(* IEC 61131-3 sources: Elmo_Master/Lasal_PRG/Elmo_EtherCAT_Test_4Axis/Class/SafetyManager (part 6) *)

      UdpReceiveData.SectionStop();
    else
      //sequence counter is not the same
      sUdpVars.WrongSequenceInResponseCnt += 1;

      //check the sequence difference, it could be a retry from other side which contains sdo data
      SequenceDifference := pConnection^.ActReceiveData.udSequenceNumber$DINT - pConnection^.ActSendData.udSequenceNumber$DINT;

      UdpReceiveData.SectionStart();
      //if Sequence difference is -1 it could be a response retry with sdo data
      if (pPacket^.Header.SdoDataLength) & (pConnection^.ActReceiveData.SdoLength = 0)
      & (pPacket^.Header.SdoDataLength <= UDP_MAX_SDO_SIZE) & (SequenceDifference = -1) then
        pConnection^.ActReceiveData.SdoLength := pPacket^.Header.SdoDataLength;
        _memcpy(ptr1:=#pConnection^.ActReceiveData.SdoData, ptr2:=#pPacket^.Data + pConnection^.ActReceiveData.PdoLength, cntr:=pConnection^.ActReceiveData.SdoLength);
      end_if;
      UdpReceiveData.SectionStop();
    end_if;

    // save safety number of other side
    pConnection^.SafetyNbrOtherSide       := pPacket^.Header.SafetyNbr;
  else
    sUdpVars.WrongReceiveUDPLength += 1;
  end_if;

END_FUNCTION

FUNCTION SafetyManager::ForwardReceivedUdpSDOs
  VAR_INPUT
    paConnections 	: ^t_aUdpConnections;
    ConnectionNo 	: UDINT;
  END_VAR
  VAR
    i               : UDINT;
    pActConnection  : ^t_UdpConnection;
    pHelpCfg        : ^t_CfgListElem;
    pHelpModule     : ^t_ModuleListElem;
    InterfaceCRC    : HDINT;
    SafetyNumber    : HDINT;
    MyPara          : CmdStruct;
    MyResult        : results;
    pDO 	          : ^SafetyCDIAS_Base::SDOHeader;
    pCompDestPath   : ^USINT;
    pHelpSafety     : ^t_SafetyComponent;
    ResponseValue   : BOOL;
    FoundTarget     : BOOL;
  END_VAR

  ResponseValue := paConnections = sUdpVars.paConnectionsToProducers;

  pActConnection := #paConnections^[0];
  for i := 0 to (ConnectionNo-1) do

    // check if there is a SDO to forward
    if pActConnection^.ActReceiveData.SdoLength then

      FoundTarget := FALSE;

      UdpReceiveData.SectionStart();

      // get a pointer to the compressed destination path
      pDO := (#pActConnection^.ActReceiveData.SdoData)$^SafetyCDIAS_Base::SDOHeader;
      if (pDO^.StdHeader.Typ.Response = ResponseValue) then
        pCompDestPath := (#pDO^.DstAdr)$^USINT;

        // check if it's addressed by topology path and it's an IP
        if ((pDO^.StdHeader.Typ AND SSDO_MASK_TYPE) = FRM_TYPECODE_SSDO_MOD_TP) & (pCompDestPath^ = INTERFACE_IP_MODE) then
          // after the mode byte we find the interface CRC
          InterfaceCRC := ((pCompDestPath + 1)$^HDINT)^;

          // search all configs, all moduleconfigs

          pHelpCfg := pConfigs;
          while pHelpCfg & pActConnection^.ActReceiveData.SdoLength do
            pHelpModule := pHelpCfg^.pFirstModuleCfg;
            while pHelpModule & pActConnection^.ActReceiveData.SdoLength do
              if pHelpModule^.ModuleInfo.InterfaceCRC = InterfaceCRC then
                // we found the interface CRC, now we have to make a connection via the SafetyNumber between the actual module config and the module handles
                pHelpSafety := pFirstSafetyComponent;
                while pHelpSafety & pActConnection^.ActReceiveData.SdoLength do
                  // we compare the safety number
                  if pHelpSafety^.SafetyNbr = pHelpModule^.ModuleInfo.SafetyNbr then

                    MyPara.uiCmd := CMD_SM_SDO_TO_MODULE;
                    MyPara.aPara[0] := pActConnection^.ActReceiveData.SdoLength;
                    MyPara.aPara[1] := (#pActConnection^.ActReceiveData.SdoData)$DINT;
                    MyPara.aPara[2] := this$DINT;

                    pHelpSafety^.pThis^.NewInst(#MyPara, #MyResult);

                    FoundTarget := TRUE;
                  end_if;

                  pHelpSafety := pHelpSafety^.pNext;
                end_while;
              end_if;

              pHelpModule := pHelpModule^.pNext;
            end_while;

            pHelpCfg := pHelpCfg^.pNext;
          end_while;
        else
          SafetyNumber := pDO^.DstAdr;

          // search by safety number and forward to internal module
          pHelpSafety := pFirstSafetyComponent;
          while pHelpSafety & pActConnection^.ActReceiveData.SdoLength do
            // we compare the safety number
            if pHelpSafety^.SafetyNbr = SafetyNumber then
              MyPara.uiCmd := CMD_SM_SDO_TO_MODULE;
              MyPara.aPara[0] := pActConnection^.ActReceiveData.SdoLength;
              MyPara.aPara[1] := (#pActConnection^.ActReceiveData.SdoData)$DINT;
              MyPara.aPara[2] := this$DINT;

              pHelpSafety^.pThis^.NewInst(#MyPara, #MyResult);

              FoundTarget := TRUE;
            end_if;

            pHelpSafety := pHelpSafety^.pNext;
          end_while;
        end_if;

        // reset length if the response bit matches (if we found it, we already forwarded it. if not, we're not going to find it next time)
        pActConnection^.ActReceiveData.SdoLength := 0;
      else
        // check which list it is
        if ResponseValue then
          sUdpVars.InvalidResponseSettingAtFowardingProducerList += 1;
        else
          sUdpVars.InvalidResponseSettingAtFowardingConsumerList += 1;
        end_if;
      end_if;

      UdpReceiveData.SectionStop();

    end_if;

    pActConnection += sizeof(t_UdpConnection);
  end_for;

END_FUNCTION

FUNCTION SafetyManager::ForwardSDO2UdpBySafetyNbr
  VAR_INPUT
    SDOLength 	: UINT;
    pSDO 	: ^USINT;
  END_VAR
  VAR_OUTPUT
    FoundTarged 	: BOOL;
  END_VAR
  VAR
    i               : UDINT;
    pActConnection  : ^t_UdpConnection;
    TargetSafetyNbr : HDINT;
    pDO 	          : ^SafetyCDIAS_Base::SDOHeader;
  END_VAR

  FoundTarged := FALSE;

  // get a pointer to the compressed destination path
  pDO := pSDO$^SafetyCDIAS_Base::SDOHeader;
  TargetSafetyNbr := pDO^.DstAdr;

  if sUdpVars.ConsumerConnectionNo then
    pActConnection := #sUdpVars.paConnectionsToConsumers^[0];
    for i := 0 to (sUdpVars.ConsumerConnectionNo-1) do
      // the safety number has to match and since it's a message to a consumer it has to be a response
      if (pActConnection^.SafetyNbrOtherSide = TargetSafetyNbr) & (pDO^.StdHeader.Typ.Response = TRUE) then
        // got it => forward the SDO
        if SDOLength <= UDP_MAX_SDO_SIZE then
          // check for unsent SDO first
          if pActConnection^.ActSendData.SdoLength = 0 then
            UdpSendData.SectionStart();

            _memcpy(ptr1:=#pActConnection^.ActSendData.SdoData, ptr2:=pSDO, cntr:=SDOLength);
            pActConnection^.ActSendData.SdoLength     := SDOLength$USINT;

            UdpSendData.SectionStop();
          else
            sUdpVars.SdoAlreadyUsedCnt += 1;
          end_if;
        else
          LogError("@046E (SafetyManager::ForwardSDO2UdpBySafetyNbr) SDO size exceeds the allowed size (Compressed Topology Path: UDP)");
        end_if;

        FoundTarged := TRUE;
        return;
      end_if;

      pActConnection += sizeof(t_UdpConnection);
    end_for;
  end_if;

  if sUdpVars.ProducerConnectionNo then
    pActConnection := #sUdpVars.paConnectionsToProducers^[0];
    for i := 0 to (sUdpVars.ProducerConnectionNo-1) do
      // the safety number has to match and since it's a message to a producer it has to be a request
      if (pActConnection^.SafetyNbrOtherSide = TargetSafetyNbr) & (pDO^.StdHeader.Typ.Response = FALSE) then
        // got it => forward the SDO
        if SDOLength <= UDP_MAX_SDO_SIZE then
          // check for unsent SDO first
          if pActConnection^.ActSendData.SdoLength = 0 then
            UdpSendData.SectionStart();

            _memcpy(ptr1:=#pActConnection^.ActSendData.SdoData, ptr2:=pSDO, cntr:=SDOLength);
            pActConnection^.ActSendData.SdoLength     := SDOLength$USINT;

            UdpSendData.SectionStop();
          else
            sUdpVars.SdoAlreadyUsedCnt += 1;
          end_if;
        else
          LogError("@046E (SafetyManager::ForwardSDO2Udp) SDO size exceeds the allowed size (Compressed Topology Path: UDP)");
        end_if;

        FoundTarged := TRUE;
        return;
      end_if;

      pActConnection += sizeof(t_UdpConnection);
    end_for;
  end_if;

END_FUNCTION

FUNCTION SafetyManager::ShareUdpConnectionInfos
  VAR
    i                 : UDINT;
    pUdpConnection    : ^t_UdpConnection;
    AnythingMissing   : BOOL;
    ActInitialized    : BOOL;
    FoundConnection   : BOOL;
    pHelpSafety       : ^t_SafetyComponent;
    pHelpCfg          : ^t_CfgListElem;
    pFSoEConnection   : ^t_FSoEConnectionDetails;
    MyPara            : CmdStruct;
    MyResult          : results;
    retcode           : iprStates;

    ModuleReadOffset  : UINT;
    ModuleReadSize    : UINT;
    ModuleWriteOffset : UINT;
    ModuleWriteSize   : UINT;
    MngReadOffset     : UINT;
    MngReadSize       : UINT;
    MngWriteOffset    : UINT;
    MngWriteSize      : UINT;
  END_VAR

  AnythingMissing := FALSE;

  if sUdpVars.ConsumerConnectionNo then
    pUdpConnection := #sUdpVars.paConnectionsToConsumers^[0];
    for i := 0 to (sUdpVars.ConsumerConnectionNo-1) do
      // check if we received something so far at this connection
      if (pUdpConnection^.ReceivedPackages & (pUdpConnection^.InfoBits.PdosInitialized = FALSE)) then
        FoundConnection := ActInitialized := FALSE;

        // check FSoE Connections in the available configs if there is a match at the interface CRC
        pHelpCfg := pConfigs;
        while pHelpCfg & (FoundConnection = FALSE) do
          pFSoEConnection := pHelpCfg^.pFirstFSoEConnection;
          while pFSoEConnection & (FoundConnection = FALSE) do
            // only interface slave connections which are not used yet are relevant
            if pFSoEConnection^.Flags.IsInterfaceConnection & (pFSoEConnection^.Flags.IsMaster = FALSE) & (pFSoEConnection^.InternalConnectionState = FCS_RESET) &
               pFSoEConnection^.pSlavePathComp & ((pFSoEConnection^.pSlavePathComp$^HDINT + 1)^ = pUdpConnection^.IFCRC) then

              // found the connection
              FoundConnection := TRUE;

              // now try to initialize it

              pHelpSafety := pFirstSafetyComponent;
              while pHelpSafety do
                if pHelpSafety^.SafetyNbr = pFSoEConnection^.OwnerSafetyNbr then
                  exit;
                end_if;

                pHelpSafety := pHelpSafety^.pNext;
              end_while;

              if pHelpSafety then
#ifdef SAFETY_DEBUG_LOGGING_ACTIVATED
#pragma message("RamAnd 20.11.2014 16:41 \ testweise mapping loggen")
                LogValue("@DBG (SafetyManager::ShareUdpConnectionInfos) <This side is Slave> ConnectionID: 0x{0}, SlaveAddress: 0x{1}, IFCRC: 0x{2}", Value:=pFSoEConnection^.ConnectionID, Value2:=pFSoEConnection^.SlaveAddress, Value3 := (pFSoEConnection^.pSlavePathComp$^HDINT + 1)^);
                LogValue("@DBG (SafetyManager::ShareUdpConnectionInfos) <This side is Slave> UdpInfo: SNr: 0x{0}, SNrOtherSide: 0x{1}, IFCRC: 0x{2}", Value:=pUdpConnection^.SafetyNbr, Value2:=pUdpConnection^.SafetyNbrOtherSide, Value3 := pUdpConnection^.IFCRC);
#endif

                // the module is slave and the managing module master
                ModuleReadOffset  := pFSoEConnection^.SlaveReadOffset;
                ModuleReadSize    := pFSoEConnection^.MasterWriteSize;
                ModuleWriteOffset := pFSoEConnection^.SlaveWriteOffset;
                ModuleWriteSize   := pFSoEConnection^.MasterReadSize;
                MngReadOffset     := 0; // offsets in managing modules are always dynamic
                MngReadSize       := pFSoEConnection^.MasterReadSize;
                MngWriteOffset    := 0; // offsets in managing modules are always dynamic
                MngWriteSize      := pFSoEConnection^.MasterWriteSize;

#ifdef SAFETY_DEBUG_LOGGING_ACTIVATED
#pragma message("RamAnd 20.11.2014 16:41 \ testweise mapping loggen")
                LogValue("@DBG (SafetyManager::ShareUdpConnectionInfos) Modul => Udp: Rd Offset Modul: 0x{0}, IP: 0x{1}, Größe: 0x{2}", Value:=ModuleReadOffset, Value2:=pUdpConnection^.IP, Value3:=ModuleReadSize);
#endif

                MyPara.uiCmd    := CMD_SM_ADD_INPUT_PDO;
                MyPara.aPara[0] := (#pUdpConnection^.ThreadSafePdoReceiveBuffer)$DINT;
                MyPara.aPara[1] := 0;
                MyPara.aPara[2] := pUdpConnection^.SafetyNbrOtherSide$DINT;
                MyPara.aPara[3] := ModuleWriteSize;
                MyPara.aPara[4] := 0;
                MyPara.aPara[5] := 0;
                MyPara.aPara[6] := 0;
                MyPara.aPara[7] := ModuleWriteOffset;
                MyPara.aPara[8] := SM_IF_VALIDITY_MARK$DINT;
                MyPara.aPara[9] := TRUE;

                retcode := pHelpSafety^.pThis^.NewInst(#MyPara, #MyResult);

                if retcode = ERROR then
                  LogError("@0848 (SafetyManager::ShareUdpConnectionInfos) Failed to add input PDO for a connection to a Consumer");

                  // mark the connection to not try again later
                  pFSoEConnection^.InternalConnectionState := FCS_NOT_INITIALIZED;

                  return;
                elsif retcode = BUSY then
                  // try again later (skip further initialisation steps)
                  return;
                end_if;

                if FSoEInputPDONo < MAX_FSOE_CONNECTIONS then
                  aFSoEInputPDOs[FSoEInputPDONo].pSafety    := pHelpSafety;
                  aFSoEInputPDOs[FSoEInputPDONo].pMem       := MyPara.aPara[0];
                  FSoEInputPDONo                            += 1;

                  pUdpConnection^.ActReceiveData.PdoLength  := ModuleWriteSize;
                else
                  LogValue("@0490 (SafetyManager::ShareUdpConnectionInfos) Maximum limit of allowed FSoE input Frames exceeded (0x{0})", Value:=MAX_FSOE_CONNECTIONS);
                  exit;
                end_if;

                if sUdpVars.ReceiveCopyCmdNo < MAX_UDP_IF_ALLOWED then
                  sUdpVars.aReceiveCopyCmds[sUdpVars.ReceiveCopyCmdNo].pSource      := (#pUdpConnection^.ActReceiveData.PdoData)$^USINT;
                  sUdpVars.aReceiveCopyCmds[sUdpVars.ReceiveCopyCmdNo].pDest        := MyPara.aPara[0]$^USINT;
                  sUdpVars.aReceiveCopyCmds[sUdpVars.ReceiveCopyCmdNo].Size         := ModuleWriteSize;
                  sUdpVars.ReceiveCopyCmdNo                                            += 1;
                else
                  LogValue("@049F (SafetyManager::ShareUdpConnectionInfos) Maximum limit of allowed UDP receive copy commands exceeded (0x{0})", Value:=MAX_UDP_IF_ALLOWED);
                  exit;
                end_if;

                MyPara.uiCmd    := CMD_SM_ADD_OUTPUT_PDO;
                MyPara.aPara[0] := 1;  // mark as interface frame PDO
                pHelpSafety^.pThis^.NewInst(#MyPara, #MyResult);

//                  pPDOElement^.SourceInfo.pPDOMem       := MyResult.aData[0]$^USINT;
//                  pPDOElement^.SourceInfo.pPDOMemDPRAM  := MyResult.aData[4]$^USINT;
//                  pPDOElement^.SourceInfo.HandlePDODPRAM:= MyResult.aData[8]$UDINT;   // Needed for Payload Support
//                  pPDOElement^.SourceInfo.OffsetPDODPRAM:= MyResult.aData[12]$UDINT;  // Needed for Payload Support

                if sUdpVars.SendCopyCmdNo < MAX_UDP_IF_ALLOWED then
                  sUdpVars.aSendCopyCmds[sUdpVars.SendCopyCmdNo].pSource      := MyResult.aData[0]$^USINT + ModuleReadOffset;
                  sUdpVars.aSendCopyCmds[sUdpVars.SendCopyCmdNo].pDest        := #pUdpConnection^.ActSendData.PdoData;
                  sUdpVars.aSendCopyCmds[sUdpVars.SendCopyCmdNo].Size         := ModuleReadSize;
                  sUdpVars.SendCopyCmdNo                                         += 1;

                  pUdpConnection^.ActSendData.PdoLength           := ModuleReadSize;
                else
                  LogValue("@049E (SafetyManager::ShareUdpConnectionInfos) Maximum limit of allowed UDP send copy commands exceeded (0x{0})", Value:=MAX_UDP_IF_ALLOWED);
                  exit;
                end_if;

#ifdef SAFETY_DEBUG_LOGGING_ACTIVATED
#pragma message("RamAnd 20.11.2014 16:41 \ testweise mapping loggen")
                LogValue("@DBG (SafetyManager::ShareUdpConnectionInfos) Udp => Modul: Wr Offset Modul: 0x{0}, IP: 0x{1}, Größe: 0x{2}", Value:=ModuleWriteOffset, Value2:=pUdpConnection^.IP, Value3:=ModuleWriteSize);
#endif

                // mark the FSoE connection as established
                pFSoEConnection^.InternalConnectionState  := FCS_CONNECTION;

                // mark the udp connection as established
                pUdpConnection^.InfoBits.PdosInitialized  := TRUE;

                // connection initialized
                ActInitialized                            := TRUE;

                // check if we have all slave addresses now
                CheckLocalSlaveAddresses();
              else
                LogValue("@495 (SafetyManager::ShareUdpConnectionInfos) Could not find safety module with safety number 0x{0} for FSoE interface connection", Value:=pFSoEConnection^.OwnerSafetyNbr);
              end_if;
            end_if;

            pFSoEConnection := pFSoEConnection^.pNext;
          end_while;

          if pHelpCfg then
            pHelpCfg := pHelpCfg^.pNext;
          end_if;
        end_while;

        if ActInitialized = FALSE then
          AnythingMissing := TRUE;
        end_if;
      elsif (pUdpConnection^.ReceivedPackages = 0) then
        AnythingMissing := TRUE;
      end_if;

      pUdpConnection += sizeof(t_UdpConnection);
    end_for;
  end_if;

  if sUdpVars.ProducerConnectionNo then
    pUdpConnection := #sUdpVars.paConnectionsToProducers^[0];
    for i := 0 to (sUdpVars.ProducerConnectionNo-1) do
      // check if we received something so far at this connection
      if (pUdpConnection^.ReceivedPackages & (pUdpConnection^.InfoBits.PdosInitialized = FALSE)) then
        FoundConnection := ActInitialized := FALSE;

        // check FSoE Connections in the available configs if there is a match at the interface CRC
        pHelpCfg := pConfigs;
        while pHelpCfg & (FoundConnection = FALSE) do
          pFSoEConnection := pHelpCfg^.pFirstFSoEConnection;
          while pFSoEConnection & (FoundConnection = FALSE) do
            // only interface master connections which are not used are relevant
            if pFSoEConnection^.Flags.IsInterfaceConnection & pFSoEConnection^.Flags.IsMaster & (pFSoEConnection^.InternalConnectionState = FCS_RESET) then
              // check if it's our connection
              if ( pFSoEConnection^.pSlavePathComp) &
                 ( pFSoEConnection^.pSlavePathComp^             = INTERFACE_IP_MODE) &
                 ((pFSoEConnection^.pSlavePathComp$^HDINT + 1)^ = pUdpConnection^.IFCRC) &
                 ((pFSoEConnection^.pSlavePathComp$^HDINT + 5)^ = pUdpConnection^.IP) then

                // found the connection
                FoundConnection := TRUE;

                // now try to initialize it

                pHelpSafety := pFirstSafetyComponent;
                while pHelpSafety do
                  if pHelpSafety^.SafetyNbr = pFSoEConnection^.OwnerSafetyNbr then
                    exit;
                  end_if;

                  pHelpSafety := pHelpSafety^.pNext;
                end_while;

                if pHelpSafety then
  #ifdef SAFETY_DEBUG_LOGGING_ACTIVATED
  #pragma message("RamAnd 20.11.2014 16:41 \ testweise mapping loggen")
                  LogValue("@DBG (SafetyManager::ShareUdpConnectionInfos) <This side is Master> ConnectionID: 0x{0}, SlaveAddress: 0x{1}, InterfaceCRC: 0x{2}", Value:=pFSoEConnection^.ConnectionID, Value2:=pFSoEConnection^.SlaveAddress, Value3 := pUdpConnection^.IFCRC);
#endif

                  // the module is master and the managing module slave
                  ModuleReadOffset  := pFSoEConnection^.MasterReadOffset;
                  ModuleReadSize    := pFSoEConnection^.MasterReadSize;
                  ModuleWriteOffset := pFSoEConnection^.MasterWriteOffset;
                  ModuleWriteSize   := pFSoEConnection^.MasterWriteSize;
                  MngReadOffset     := 0; // offsets in managing modules are always dynamic
                  MngReadSize       := pFSoEConnection^.MasterWriteSize;
                  MngWriteOffset    := 0; // offsets in managing modules are always dynamic
                  MngWriteSize      := pFSoEConnection^.MasterReadSize;

  #ifdef SAFETY_DEBUG_LOGGING_ACTIVATED
  #pragma message("RamAnd 20.11.2014 16:41 \ testweise mapping loggen")
                  LogValue("@DBG (SafetyManager::ShareUdpConnectionInfos) Modul => Udp: Rd Offset Modul: 0x{0}, IP: 0x{1}, Größe: 0x{2}", Value:=ModuleReadOffset, Value2:=pUdpConnection^.IP, Value3:=ModuleReadSize);
  #endif

                  MyPara.uiCmd    := CMD_SM_ADD_INPUT_PDO;
                  MyPara.aPara[0] := (#pUdpConnection^.ThreadSafePdoReceiveBuffer)$DINT;
                  MyPara.aPara[1] := 0;
                  MyPara.aPara[2] := pUdpConnection^.SafetyNbrOtherSide$DINT;
                  MyPara.aPara[3] := ModuleWriteSize;
                  MyPara.aPara[4] := 0;
                  MyPara.aPara[5] := 0;
                  MyPara.aPara[6] := 0;
                  MyPara.aPara[7] := ModuleWriteOffset;
                  MyPara.aPara[8] := SM_IF_VALIDITY_MARK$DINT;
                  MyPara.aPara[9] := TRUE;

                  retcode := pHelpSafety^.pThis^.NewInst(#MyPara, #MyResult);

                  if retcode = ERROR then
                    LogError("@0849 (SafetyManager::ShareUdpConnectionInfos) Failed to add input PDO for a connection to a Producer");

                    // mark the connection to not try again later
                    pFSoEConnection^.InternalConnectionState := FCS_NOT_INITIALIZED;

                    return;
                  elsif retcode = BUSY then
                    // try again later (skip further initialisation steps)
                    return;
                  end_if;

                  if FSoEInputPDONo < MAX_FSOE_CONNECTIONS then
                    aFSoEInputPDOs[FSoEInputPDONo].pSafety    := pHelpSafety;
                    aFSoEInputPDOs[FSoEInputPDONo].pMem       := MyPara.aPara[0];
                    FSoEInputPDONo += 1;

                    pUdpConnection^.ActReceiveData.PdoLength  := ModuleWriteSize;
                  else
                    LogValue("@0490 (SafetyManager::ShareUdpConnectionInfos) Maximum limit of allowed FSoE input Frames exceeded (0x{0})", Value:=MAX_FSOE_CONNECTIONS);
                    exit;
                  end_if;

                  if sUdpVars.ReceiveCopyCmdNo < MAX_UDP_IF_ALLOWED then
                    sUdpVars.aReceiveCopyCmds[sUdpVars.ReceiveCopyCmdNo].pSource  := (#pUdpConnection^.ActReceiveData.PdoData)$^USINT;
                    sUdpVars.aReceiveCopyCmds[sUdpVars.ReceiveCopyCmdNo].pDest    := MyPara.aPara[0]$^USINT;
                    sUdpVars.aReceiveCopyCmds[sUdpVars.ReceiveCopyCmdNo].Size     := ModuleWriteSize;
                    sUdpVars.ReceiveCopyCmdNo                                        += 1;
                  else
                    LogValue("@049F (SafetyManager::ShareUdpConnectionInfos) Maximum limit of allowed UDP receive copy commands exceeded (0x{0})", Value:=MAX_UDP_IF_ALLOWED);
                    exit;
                  end_if;

                  MyPara.uiCmd      := CMD_SM_ADD_OUTPUT_PDO;
                  MyPara.aPara[0]   := 1;  // mark as interface frame PDO
                  pHelpSafety^.pThis^.NewInst(#MyPara, #MyResult);

  //                  pPDOElement^.SourceInfo.pPDOMem       := MyResult.aData[0]$^USINT;
  //                  pPDOElement^.SourceInfo.pPDOMemDPRAM  := MyResult.aData[4]$^USINT;
  //                  pPDOElement^.SourceInfo.HandlePDODPRAM:= MyResult.aData[8]$UDINT;   // Needed for Payload Support
  //                  pPDOElement^.SourceInfo.OffsetPDODPRAM:= MyResult.aData[12]$UDINT;  // Needed for Payload Support

                  if sUdpVars.SendCopyCmdNo < MAX_UDP_IF_ALLOWED then
                    sUdpVars.aSendCopyCmds[sUdpVars.SendCopyCmdNo].pSource      := MyResult.aData[0]$^USINT + ModuleReadOffset;
                    sUdpVars.aSendCopyCmds[sUdpVars.SendCopyCmdNo].pDest        := #pUdpConnection^.ActSendData.PdoData;
                    sUdpVars.aSendCopyCmds[sUdpVars.SendCopyCmdNo].Size         := ModuleReadSize;
                    sUdpVars.SendCopyCmdNo                                         += 1;

                    pUdpConnection^.ActSendData.PdoLength                             := ModuleReadSize;
                  else
                    LogValue("@049E (SafetyManager::ShareUdpConnectionInfos) Maximum limit of allowed UDP send copy commands exceeded (0x{0})", Value:=MAX_UDP_IF_ALLOWED);
                    exit;
                  end_if;

  #ifdef SAFETY_DEBUG_LOGGING_ACTIVATED
  #pragma message("RamAnd 20.11.2014 16:41 \ testweise mapping loggen")
                  LogValue("@DBG (SafetyManager::ShareUdpConnectionInfos) Udp => Modul: Wr Offset Modul: 0x{0}, IP: 0x{1}, Größe: 0x{2}", Value:=ModuleWriteOffset, Value2:=pUdpConnection^.IP, Value3:=ModuleWriteSize);
  #endif

                  // mark the FSoE connection as established
                  pFSoEConnection^.InternalConnectionState  := FCS_CONNECTION;

                  // mark the udp connection as established
                  pUdpConnection^.InfoBits.PdosInitialized  := TRUE;

                  // connection initialized
                  ActInitialized                            := TRUE;

                  // check if we have all slave addresses now
                  CheckLocalSlaveAddresses();
                else
                  LogValue("@0495 (SafetyManager::ShareUdpConnectionInfos) Could not find safety module with safety number 0x{0} for FSoE interface connection", Value:=pFSoEConnection^.OwnerSafetyNbr);
                end_if;

              end_if;

            end_if;

            pFSoEConnection := pFSoEConnection^.pNext;
          end_while;

          pHelpCfg := pHelpCfg^.pNext;
       end_while;

        if ActInitialized = FALSE then
          AnythingMissing := TRUE;
        end_if;
      elsif (pUdpConnection^.ReceivedPackages = 0) then
        AnythingMissing := TRUE;
      end_if;

      pUdpConnection += sizeof(t_UdpConnection);
    end_for;
  end_if;

  // if all available udp connections are initialized => set the marker for not coming here any more
  if AnythingMissing = FALSE then
    sUdpVars.ConnectionsInitialized := TRUE;

    // update scheduler grid
    SetUdpSchedulerGrid();
  end_if;

END_FUNCTION

FUNCTION SafetyManager::SetUdpSchedulerGrid
  VAR
    Temp            : UDINT;
    bGetRequestTimeout : BOOL;
  END_VAR

  bGetRequestTimeout := FALSE;

  // we can only calculate if there are producer connections => otherwise the scheduler is not active
  if sUdpVars.ProducerConnectionNo then

    // the timeout is calculated so we could fit 4 timed out transmissions into the watchdog time (watchdog = 2*transmission time)
    Temp := sUdpVars.LowestTransmissionTime_ms * 2 / 4;

    // if the result is smaller than the minimum timeout => set it to the minimum
    if Temp < UDP_MIN_REQUEST_TIMEOUT then
      Temp := UDP_MIN_REQUEST_TIMEOUT;
    end_if;

    sUdpVars.CalculatedRequestTimeout := Temp;
    bGetRequestTimeout := TRUE;
  else
    // activate the default settings (min settings)
    sUdpVars.CalculatedRequestTimeout := UDP_MIN_REQUEST_TIMEOUT;
  end_if;

  // use default value for request time
  sUdpVars.CalculatedRequestTime    := UDP_MIN_REQUEST_TIME;

  //check for advanced request time from user
  if sUdpVars.udAdvancedRequestCycle >= UDP_MIN_REQUEST_TIME
  & sUdpVars.udAdvancedRequestCycle <= (sUdpVars.CalculatedRequestTimeout/2)  then
    sUdpVars.CalculatedRequestTime := sUdpVars.udAdvancedRequestCycle;
  else
    //only log error if we got calculated request timeout and value is not zero
    if bGetRequestTimeout = TRUE & sUdpVars.udAdvancedResponseTimeout <> 0 & bd_SingleLog.SetUdpRequestCycleFailed = FALSE then
      LogValue("@04D6 (SafetyManager::SetUdpSchedulerGrid) [SL] The value of 0x{0} for the UDP Request Cycle is not valid! The maximum value is 0x{1}", Value:=sUdpVars.udAdvancedRequestCycle, (sUdpVars.CalculatedRequestTimeout/2));
      bd_SingleLog.SetUdpRequestCycleFailed := TRUE;
    end_if;
  end_if;

  // always use the min settings for the responses
  sUdpVars.CalculatedResponseTime    := UDP_MIN_RESPONSE_TIME;
  sUdpVars.CalculatedResponseTimeout := UDP_MIN_RESPONSE_TIMEOUT;

  //check for advanced response timeout from user
  if sUdpVars.udAdvancedResponseTimeout >= UDP_MIN_RESPONSE_TIMEOUT then
    sUdpVars.CalculatedResponseTimeout := sUdpVars.udAdvancedResponseTimeout;
  else
    // only log error if value is not zero
    if sUdpVars.udAdvancedResponseTimeout <> 0 & bd_SingleLog.SetUdpResponseTimeoutFailed = FALSE then
      LogValue("@04D7 (SafetyManager::SetUdpSchedulerGrid) [SL] The value of 0x{0} for the UDP Response Timeout is not valid! The minimum value is 0x{1}", Value:=sUdpVars.udAdvancedResponseTimeout, UDP_MIN_RESPONSE_TIMEOUT);
      bd_SingleLog.SetUdpResponseTimeoutFailed := TRUE;
    end_if;
  end_if;

  // if the override values are set => activate them here to override all other settings
  if sUdpVars.udOverrideCycleTime then
    // set the scheduler grid for requests and resonses according to the override value
    sUdpVars.CalculatedRequestTime  := sUdpVars.udOverrideCycleTime;
    sUdpVars.CalculatedResponseTime := sUdpVars.udOverrideCycleTime;
  end_if;

  if sUdpVars.udOverrideTimeout then
    // set the timeout value for requests and resonses according to the override value
    sUdpVars.CalculatedRequestTimeout  := sUdpVars.udOverrideTimeout;
    sUdpVars.CalculatedResponseTimeout := sUdpVars.udOverrideTimeout;
  end_if;

END_FUNCTION

FUNCTION SafetyManager::UdpResponseScheduler
  VAR
    pActResponseEntry : ^t_UdpConnection;
    pActRetryEntry    : ^t_UdpConnection;
    tmpretcode        : DINT;
    i                 : UDINT;
  END_VAR

  //point to actual request-entry
  pActResponseEntry := #sUdpVars.paConnectionsToConsumers^[sUdpVars.ResponseScheduler.ActRequestedIndex];

  //send a request every TRequestTime x Cycnt Cycle
  if ((sUdpVars.ResponseScheduler.CyCnt MOD sUdpVars.CalculatedResponseTime) = 0) then

    // search through the list if something has to be sent (check also for changes in the data)
    for i := 0 to sUdpVars.ConsumerConnectionNo-1 do

      //only send a request if not waiting for a response and the IP is valid (on cleaning out the connections some may be set to 0)
      if (pActResponseEntry^.WaitForResponse = FALSE) & (pActResponseEntry^.IP <> 0) & (pActResponseEntry^.SendResponse = TRUE) then

        //send request to mover of actual entry
        tmpretcode := SendUdpResponse(pActResponseEntry);
        if tmpretcode >= 0 then

          //if sending was successful we are waiting for a response
          pActResponseEntry^.WaitForResponse := TRUE;
          pActResponseEntry^.SendResponse    := FALSE;
          pActResponseEntry^.TLastRequest      := ops.tAbsolute;
          pActResponseEntry^.RequestRetries    := 0;

        else
          //unable to send request
          if bd_SingleLog.SendUdpRspFailed = FALSE then
            bd_SingleLog.SendUdpRspFailed := TRUE;
            LogError("@04A0 (SafetyManager::UdpResponseScheduler) [SL] Failed to send udp response");
          end_if;
        end_if;

      end_if;

      //increase actual index
      if sUdpVars.ResponseScheduler.ActRequestedIndex < (sUdpVars.ConsumerConnectionNo-1) then
        sUdpVars.ResponseScheduler.ActRequestedIndex += 1;
      else
        //when reaching last entry -> reset index
        sUdpVars.ResponseScheduler.ActRequestedIndex := 0;
      end_if;

      pActResponseEntry := #sUdpVars.paConnectionsToConsumers^[sUdpVars.ResponseScheduler.ActRequestedIndex];
    end_for;

  // between the normal requests we do the retries
  elsif ((sUdpVars.ResponseScheduler.CyCnt MOD UDP_RETRY_TIME) = 0) then

    pActRetryEntry := #sUdpVars.paConnectionsToConsumers^[0];

    // check if we have to send a retry
    for i := 0 to sUdpVars.ConsumerConnectionNo-1 do

      // look if we actual wait for a response to send retries and check if we didn't receive data in time
      if (pActRetryEntry^.WaitForResponse = TRUE) & ((ops.tAbsolute - pActRetryEntry^.TLastRequest) > sUdpVars.CalculatedResponseTimeout) then

        if pActRetryEntry^.RequestRetries >= UDP_MAX_RETRIES then

          pActRetryEntry^.MaxRetryCnt          += 1;
          pActRetryEntry^.WaitForResponse      := FALSE;
          //don't reset flag here, because it's possible we receive an old sequence counter with next package, which leads to an error at FSoE communication
          //pActRetryEntry^.bSequenceCntReceived := FALSE; //reset flag to allow sequence counter for new udp communication

        // only if the IP is valid
        elsif (pActRetryEntry^.IP <> 0) then

          //send retry to actual cpu
          tmpretcode := SendUdpResponse(pActRetryEntry);
          if tmpretcode >= 0 then
            pActRetryEntry^.TLastRequest   := ops.tAbsolute;
            pActRetryEntry^.RequestRetries += 1;
            exit;
          else
            //unable to send retry
            if bd_SingleLog.SendUdpRspRetryFailed = FALSE then
              bd_SingleLog.SendUdpRspRetryFailed := TRUE;
              LogError("@049D (SafetyManager::UdpResponseScheduler) [SL] Failed to send udp retry");
            end_if;
          end_if;
        end_if;

      end_if;

      pActRetryEntry += sizeof(t_UdpConnection);

    end_for;

  end_if;

  sUdpVars.ResponseScheduler.CyCnt += 1;

END_FUNCTION

FUNCTION SafetyManager::SendUdpResponse
  VAR_INPUT
    pConnection 	: ^t_UdpConnection;
  END_VAR
  VAR_OUTPUT
    retcode 	: DINT;
  END_VAR
  VAR
    udActSendLength : UDINT;
  END_VAR

  sUdpVars.pTempSendBufferCy^.Header.Command   := t_UdpCommand::UdpCmd_DataRsp;
  //The current header version is set here so that the other side knows which version is supported.
  sUdpVars.pTempSendBufferCy^.Header.State     := t_UdpPacketHeaderV2.State.IsFromProducer + UDP_HEADER_ACTVERSION;
  sUdpVars.pTempSendBufferCy^.Header.IFCRC     := pConnection^.IFCRC;
  sUdpVars.pTempSendBufferCy^.Header.SafetyNbr := pConnection^.SafetyNbr;

  UdpSendData.SectionStart();

  //check for new header version with extended sequence number (4Byte)
  if pConnection^.ActSendData.usHeaderVersion >= UDP_HEADER_VERSION_V2 then

    sUdpVars.pTempSendBufferCy^.Header.SequenceNumber := pConnection^.ActSendData.udSequenceNumber;

    udActSendLength := sizeof(t_UdpPacketHeaderV2);

    if pConnection^.ActSendData.PdoLength then
      sUdpVars.pTempSendBufferCy^.Header.PdoDataLength  := pConnection^.ActSendData.PdoLength;
      _memcpy(ptr1:=#sUdpVars.pTempSendBufferCy^.Data, ptr2:=#pConnection^.ActSendData.PdoData, cntr:=pConnection^.ActSendData.PdoLength);
      udActSendLength += pConnection^.ActSendData.PdoLength;
    else
      sUdpVars.pTempSendBufferCy^.Header.PdoDataLength  := 0;
    end_if;

    if pConnection^.ActSendData.SdoLength then
      sUdpVars.pTempSendBufferCy^.Header.SdoDataLength  := pConnection^.ActSendData.SdoLength;
      _memcpy(ptr1:=#sUdpVars.pTempSendBufferCy^.Data + pConnection^.ActSendData.PdoLength, ptr2:=#pConnection^.ActSendData.SdoData, cntr:=pConnection^.ActSendData.SdoLength);
      udActSendLength += pConnection^.ActSendData.SdoLength;
    else
      sUdpVars.pTempSendBufferCy^.Header.SdoDataLength  := 0;
    end_if;
  else
    //use old headerversion with 1byte Sequence Counter
    sUdpVars.pTempSendBufferCy^$t_UdpPacketV1.Header.SequenceNumber := pConnection^.ActSendData.usSequenceNumber;

    udActSendLength := sizeof(t_UdpPacketHeaderV1);

    if pConnection^.ActSendData.PdoLength then
      sUdpVars.pTempSendBufferCy^$t_UdpPacketV1.Header.PdoDataLength  := pConnection^.ActSendData.PdoLength;
      _memcpy(ptr1:=#sUdpVars.pTempSendBufferCy^$t_UdpPacketV1.Data, ptr2:=#pConnection^.ActSendData.PdoData, cntr:=pConnection^.ActSendData.PdoLength);
      udActSendLength += pConnection^.ActSendData.PdoLength;
    else
      sUdpVars.pTempSendBufferCy^$t_UdpPacketV1.Header.PdoDataLength  := 0;
    end_if;

    if pConnection^.ActSendData.SdoLength then
      sUdpVars.pTempSendBufferCy^$t_UdpPacketV1.Header.SdoDataLength  := pConnection^.ActSendData.SdoLength;
      _memcpy(ptr1:=#sUdpVars.pTempSendBufferCy^$t_UdpPacketV1.Data + pConnection^.ActSendData.PdoLength, ptr2:=#pConnection^.ActSendData.SdoData, cntr:=pConnection^.ActSendData.SdoLength);
      udActSendLength += pConnection^.ActSendData.SdoLength;
    else
      sUdpVars.pTempSendBufferCy^$t_UdpPacketV1.Header.SdoDataLength  := 0;
    end_if;

  end_if;

  UdpSendData.SectionStop();

  retcode := SendUDPData(sUdpVars.pTempSendBufferCy, udActSendLength, pConnection^.IP);

  sUdpVars.SendCnt += 1;

  if retcode < 0 then
    // error at sending
    sUdpVars.LastSendError := retcode;
    sUdpVars.SendErrorCnt += 1;
  else
    // only valid one-time
    pConnection^.ActSendData.SdoLength    := 0;

    pConnection^.SentPackages += 1;
  end_if;

END_FUNCTION

FUNCTION SafetyManager::UdpTask

  while TRUE do

        // if there is no error and we got UDP stuff going on => do it
    if (sUdpVars.ProducerConnectionNo | ((sUdpVars.UdpInit AND 2#11) = (t_UdpInit.FSoEAvailable OR t_UdpInit.ProvidesIF))) then
      if sUdpVars.UdpInit.CallBackInstalled = FALSE then

        //add callback info for receiving udp packages
        AddCallBackInfo(this, #ReceiveUDPData());

        sUdpVars.UdpInit.CallBackInstalled := TRUE;
      end_if;

      SafetyUDP::CyWork(0);

      // no SDOs or scheduling when we reinitialize
      if CommInitialized & (InitSSW > _ClearRoutingInfos) then
        // check initialisation of the connections
        if (sUdpVars.ConnectionsInitialized = FALSE) & ((LastUdpIfCfgDistribution = 0) | ((ops.tAbsolute - LastUdpIfCfgDistribution) > SM_INTERFACE_CONFIG_SEND_PAUSE)) then

          ShareUdpConnectionInfos();

          // remember when the config has been distributed, to not spam the other sides
          LastUdpIfCfgDistribution := ops.tAbsolute;
        end_if;

        // only if we're a consumer and have producers to contact
        if sUdpVars.ProducerConnectionNo then

          // work the connections (send requests)
          UdpRequestScheduler();

          // forward the SDOs from the producer (responses)
          ForwardReceivedUdpSDOs(paConnections:=sUdpVars.paConnectionsToProducers, ConnectionNo:=sUdpVars.ProducerConnectionNo);
        end_if;

        // if there are consumers, we may distribute new SDO data
        if sUdpVars.ConsumerConnectionNo then

          // work the connections (send responses)
          UdpResponseScheduler();

          // forward the SDOs from the consumers (requests)
          ForwardReceivedUdpSDOs(paConnections:=sUdpVars.paConnectionsToConsumers, ConnectionNo:=sUdpVars.ConsumerConnectionNo);
        end_if;
      end_if;
    end_if;

    To_MultiTask.TASKDELAY(timeout0:=1);
  end_while;

END_FUNCTION

FUNCTION SafetyManager::TimeSyncModuleAvailable
  VAR_INPUT
    pTimeSyncElement 	: ^t_TimeSyncElement;
  END_VAR
  VAR_OUTPUT
    Available 	: BOOL;
  END_VAR

  if pTimeSyncElement^.InfoBits.IsMissingOptional | (pTimeSyncElement^.pSafety & (pTimeSyncElement^.pSafety^.SafetyNbr = 0)) then
    Available := FALSE;
  else
    Available := TRUE;
  end_if;

END_FUNCTION

FUNCTION SafetyManager::ReinitEverything
  VAR
    MyPara 	  : CmdStruct;
    MyResult 	: results;
  END_VAR

  // new safety project detected (different crc) => reinit the system (similar to disconnect)
  MyPara.uiCmd := CMD_SM_DISCONNECT;
  MyPara.aPara[0] := 0; // set length of further parameters to 0
// don't disconnect connected managing modules. if there is any difference in the communication, it will be interchanged via special SDO frames (CMD_SM_IF_MODULE_INFO...)
//  TellAllInterfaceManagingModules(#MyPara, #MyResult);
  TellAllSafetyModules(#MyPara, #MyResult);             // tell all of our local safety modules that there's a new config => reinitialize

  ClassState := 0;

  // reset module sync no (no more modules synchron)
  ModuleSyncNo := 0;

  // restart initialisation (maybe we had no clue about interfaceframes when initialising the first time)
  InitSSW := _ClearRoutingInfos;

END_FUNCTION

FUNCTION SafetyManager::CheckCustomConnectionValid
  VAR_INPUT
    pConnection 	: ^t_FSoEConnectionDetails;
    pIFFSoEInfo 	: ^t_FSoEConnInfo;
  END_VAR
  VAR_OUTPUT
    bIsCustomConnValid 	: BOOL;
  END_VAR

  // This method checks if the passed connection and FSoE Interface are a Valid custom connection
  // This check replaces the slave address check for normal FSoE Interface frames. (s. FinalizePDOMapping)
  // (The slave addresses may not valid for custom connections at this point)

  bIsCustomConnValid := FALSE;

  if pConnection = NIL | pIFFSoEInfo = NIL | pIFFSoEInfo^.pManaging = NIL then
    return;
  end_if;

  if pConnection^.Flags.IsMaster then

    // Check for custom ip address in compressed path
    // Check for HWT_ESCAPE_SAFETY_CUSTOM in uncompressed path
    // pConnection^.pSlavePathComp: 1 Byte Type, 4 Byte IF CRC, 4 Byte Custom IP Addr,
    // example : 03 59 8C AE 3D 00 00 00 02 FF FF FF
    // pIFFSoEInfo^.pManaging^.pModulePath: 2 Byte Length, 1 Byte Domain No, 1 Byte Escape Sequence, 1 Byte Custom IP Addr
    // example : 03 00 00 8A 02
    if pConnection^.pSlavePathComp & pConnection^.SlavePathCompLen > 8 &                    // Pointer + length (Custom IP = Byte 9)
       (pConnection^.pSlavePathComp^ = 3) &                                                 // Type Code
       pIFFSoEInfo^.pManaging^.pModulePath & (pIFFSoEInfo^.pManaging^.pModulePath^ >= 3) &  // Pointer + length
       ((pConnection^.pSlavePathComp+5)^$UDINT AND 16#00FFFFFF) = 0 &                       // Custom IP
       (pIFFSoEInfo^.pManaging^.pModulePath+3)^ = HWT_ESCAPE_SAFETY_CUSTOM  then            // Escape Sequence
      // Compare Custom IDs
      if (pConnection^.pSlavePathComp + 8)^ = (pIFFSoEInfo^.pManaging^.pModulePath+4)^ then
        bIsCustomConnValid := TRUE;
      end_if;

    end_if;

  else

    // Check IFCRC in compressed path
    // Check for HWT_ESCAPE_SAFETY_CUSTOM in uncompressed path
    // pConnection^.pSlavePathComp: 1 Byte Type, 4 Byte IF CRC
    // example : 03 59 8C AE 3D FF FF FF
    // pIFFSoEInfo^.pManaging^.pModulePath: 2 Byte Length, 1 Byte Domain No, 1 Byte Escape Sequence, 1 Byte Custom IP Addr
    // example : 03 00 00 8A 02
    if pConnection^.pSlavePathComp & pConnection^.SlavePathCompLen > 5 &                    // Pointer + length (IFCRC = Byte 1, 4Byte CRC Data )
       (pConnection^.pSlavePathComp^ = 3) &                                                 // Type Code
       pIFFSoEInfo^.pManaging^.pModulePath & (pIFFSoEInfo^.pManaging^.pModulePath^ >= 3) &  // Pointer + length
       (pIFFSoEInfo^.pManaging^.pModulePath+3)^ = HWT_ESCAPE_SAFETY_CUSTOM then             // Escape Sequence

      // Compare IFCRC (Cannot compare Custom IDs because (pConnection^.pSlavePathComp + 8)^ may not be valid yet at this time
      if (pConnection^.pSlavePathComp+1)^$UDINT = pIFFSoEInfo^.FromOtherSide.InterfaceCRC then
        bIsCustomConnValid := TRUE;
      end_if;

    end_if;

  end_if;

END_FUNCTION

FUNCTION SafetyManager::ShareSingleConnectionInfos
	VAR_INPUT
		pMasterConnection 	: ^t_FSoEConnectionDetails;
		pModuleConfig 	: ^t_ModuleListElem;
	END_VAR
  VAR
  	pMasterModuleCfg  : ^t_ModuleListElem;
  	pSlaveModuleCfg   : ^t_ModuleListElem;
    pActModuleCfg     : ^t_ModuleListElem;
    pHelpSafety       : ^t_SafetyComponent;
    pMasterSafety     : ^t_SafetyComponent;
    pSlaveSafety      : ^t_SafetyComponent;
    MyPara 	          : CmdStruct;
    MyResult	        : results;
    pPDOReadData      : pVoid;
    i                 : UDINT;
    IsInList          : BOOL;
  END_VAR

//*****************************************************************************
//** TELL THE MODULES WHAT DATA TO COPY IN REALTIME                          **
//*****************************************************************************

  // get the master and slave module configuration of this connection

  // master module configuration is always the first one in the list
  pMasterModuleCfg  := pModuleConfig;

  // search for the slave config via the path stored in the connection
  pSlaveModuleCfg   := NIL;
  pActModuleCfg     := pModuleConfig;

  if pMasterConnection^.Flags.HWPathIsFSoEAddr = 0 then // Do not check in this case because Slave Module does not exist in the SCP configuration

    while pActModuleCfg do
      if (pActModuleCfg^.ModuleInfo.pPath^ = pMasterConnection^.pSlavePath^) &
         (To_StdLib.MemCmp(pActModuleCfg^.ModuleInfo.pPath+1, pMasterConnection^.pSlavePath+1, pMasterConnection^.pSlavePath^+1) = 0) then

        pSlaveModuleCfg := pActModuleCfg;
        exit;
      end_if;

      pActModuleCfg := pActModuleCfg^.pNext;
    end_while;

    if pSlaveModuleCfg = NIL then
      return;
    end_if;
  end_if;

  // get the object this pointers via the hardware paths
  pMasterSafety := NIL;
  pSlaveSafety  := NIL;

  // Search for Master Object
  pHelpSafety := pFirstSafetyComponent;
  while pHelpSafety do
    if pHelpSafety^.PathLen &
       (pMasterModuleCfg^.ModuleInfo.pPath^ = pHelpSafety^.pPath^) &
       (To_StdLib.MemCmp(pHelpSafety^.pPath + 1, pMasterModuleCfg^.ModuleInfo.pPath + 2, pHelpSafety^.pPath^) = 0) then
      pMasterSafety := pHelpSafety;
      exit;
    else
      pHelpSafety := pHelpSafety^.pNext;
    end_if;
  end_while;

  // Search for Slave Object
  pHelpSafety := pFirstSafetyComponent;
  if pMasterConnection^.Flags.HWPathIsFSoEAddr = 0 then // Do not check pSlaveModuleCfg this case because Slave Module does not exist in the SCP configuration
    while pHelpSafety do
      if pHelpSafety^.PathLen &
         (pSlaveModuleCfg^.ModuleInfo.pPath^ = pHelpSafety^.pPath^) &
         (To_StdLib.MemCmp(pHelpSafety^.pPath + 1, pSlaveModuleCfg^.ModuleInfo.pPath + 2, pHelpSafety^.pPath^) = 0) then
        pSlaveSafety := pHelpSafety;
        exit;
      else
        pHelpSafety := pHelpSafety^.pNext;
      end_if;
    end_while;
  else
    while pHelpSafety do
      if pHelpSafety^.PathLen &
         (pMasterConnection^.pSlavePath^ = pHelpSafety^.pPath^) &
         (To_StdLib.MemCmp(pHelpSafety^.pPath + 1, pMasterConnection^.pSlavePath + 2, pHelpSafety^.pPath^) = 0) then
        pSlaveSafety := pHelpSafety;
        exit;
      else
        pHelpSafety := pHelpSafety^.pNext;
      end_if;
    end_while;
  end_if;

  if pMasterSafety & pSlaveSafety then

    // we start with the safe outputs: get the data pointer from the master and give it to the slave
    MyPara.uiCmd    := CMD_SM_ADD_OUTPUT_PDO;
    MyResult.uiLng  := 0;
    pMasterSafety^.pThis^.NewInst(#MyPara, #MyResult);

    if MyResult.uiLng <> 4 then
      LogError("@048F (SafetyManager::ShareSingleConnectionInfos) Invalid return value when asking the master safety module for it's pointer to the PDO read data!");
      return;
    end_if;

    pPDOReadData := MyResult.aData[0]$pVoid;

  #ifdef SAFETY_DEBUG_LOGGING_ACTIVATED
  #pragma message("RamAnd 20.11.2014 16:41 \ testweise mapping loggen")
    LogValue("@DBG (SafetyManager::ShareSingleConnectionInfos) ConnectionID: {0}, SlaveAddress: {1}", Value:=pMasterConnection^.ConnectionID, Value2:=pMasterConnection^.SlaveAddress);
    LogValue("@DBG (SafetyManager::ShareSingleConnectionInfos) MasterSafetyNbr: {0}, SlaveSafetyNbr: {1}", Value:=pMasterSafety^.SafetyNbr, Value2:=pSlaveSafety^.SafetyNbr);
    LogValue("@DBG (SafetyManager::ShareSingleConnectionInfos) MasterReadOffset: {0}, MasterReadSize: {1}, SlaveWriteOffset: {2}", Value:=pMasterConnection^.MasterReadOffset, Value2:=pMasterConnection^.MasterReadSize, Value3 := pMasterConnection^.SlaveWriteOffset);
  #endif

    // check if it's in the list
    IsInList := FALSE;
    if FSoEInputPDONo then
      for i := 0 to (FSoEInputPDONo-1) do
        if ((aFSoEInputPDOs[i].pSafety = pSlaveSafety)  & (aFSoEInputPDOs[i].pMem = pPDOReadData$DINT + pMasterConnection^.MasterReadOffset)) then
          aFSoEInputPDOs[FSoEInputPDONo].pSafety    := pMasterSafety;
          aFSoEInputPDOs[FSoEInputPDONo].pMem       := MyPara.aPara[0];
          IsInList := TRUE;
        end_if;
      end_for;
    end_if;

    if IsInList = FALSE then
      MyPara.uiCmd    := CMD_SM_ADD_INPUT_PDO;
      MyPara.aPara[0] := pPDOReadData$DINT + pMasterConnection^.MasterReadOffset;
      MyPara.aPara[2] := pMasterConnection^.OwnerSafetyNbr$DINT;
      MyPara.aPara[3] := pMasterConnection^.MasterReadSize;
      MyPara.aPara[4] := pMasterSafety^.InfoBits.IsOptional;
      MyPara.aPara[7] := pMasterConnection^.SlaveWriteOffset;
      MyPara.aPara[8] := SM_IF_VALIDITY_MARK$DINT;
      MyPara.aPara[9] := pMasterConnection^.Flags.IsInterfaceConnection;
      pSlaveSafety^.pThis^.NewInst(#MyPara, #MyResult);

      if FSoEInputPDONo < MAX_FSOE_CONNECTIONS then
        aFSoEInputPDOs[FSoEInputPDONo].pSafety    := pSlaveSafety;
        aFSoEInputPDOs[FSoEInputPDONo].pMem       := MyPara.aPara[0];
        FSoEInputPDONo += 1;
      else
        LogValue("@0490 (SafetyManager::ShareSingleConnectionInfos) Maximum limit of allowed FSoE input Frames exceeded (0x{0})", Value:=MAX_FSOE_CONNECTIONS);
      end_if;
    end_if;

    // safe inputs: get the data pointer from the slave and give it to the master
    MyPara.uiCmd    := CMD_SM_ADD_OUTPUT_PDO;
    MyResult.uiLng  := 0;
    pSlaveSafety^.pThis^.NewInst(#MyPara, #MyResult);

    if MyResult.uiLng <> 4 then
      LogError("@0491 (SafetyManager::ShareSingleConnectionInfos) Invalid return value when asking the slave safety module for it's pointer to the PDO read data!");
      return;
    end_if;

    pPDOReadData := MyResult.aData[0]$pVoid;

  #ifdef SAFETY_DEBUG_LOGGING_ACTIVATED
  #pragma message("RamAnd 20.11.2014 16:41 \ testweise mapping loggen")
    LogValue("@DBG (SafetyManager::ShareSingleConnectionInfos) SlaveReadOffset: {0}, SlaveReadSize: {1}, MasterWriteOffset: {2}", Value:=pMasterConnection^.SlaveReadOffset, Value2:=pMasterConnection^.MasterWriteSize, Value3 := pMasterConnection^.MasterWriteOffset);
  #endif

    // check if it's in the list
    IsInList := FALSE;
    if FSoEInputPDONo then
      for i := 0 to (FSoEInputPDONo-1) do
        if ((aFSoEInputPDOs[i].pSafety = pMasterSafety)  & (aFSoEInputPDOs[i].pMem = pPDOReadData$DINT + pMasterConnection^.SlaveReadOffset)) then
          aFSoEInputPDOs[FSoEInputPDONo].pSafety    := pMasterSafety;
          aFSoEInputPDOs[FSoEInputPDONo].pMem       := MyPara.aPara[0];
          IsInList := TRUE;
        end_if;
      end_for;
    end_if;

    if IsInList = FALSE then

      MyPara.uiCmd    := CMD_SM_ADD_INPUT_PDO;
      MyPara.aPara[0] := pPDOReadData$DINT + pMasterConnection^.SlaveReadOffset;
      MyPara.aPara[2] := pSlaveSafety^.SafetyNbr$DINT;
      MyPara.aPara[3] := pMasterConnection^.MasterWriteSize;
      MyPara.aPara[4] := pSlaveSafety^.InfoBits.IsOptional;
      MyPara.aPara[7] := pMasterConnection^.MasterWriteOffset;
      MyPara.aPara[8] := 0;
      MyPara.aPara[9] := 0;
      pMasterSafety^.pThis^.NewInst(#MyPara, #MyResult);

      if FSoEInputPDONo < MAX_FSOE_CONNECTIONS then
        aFSoEInputPDOs[FSoEInputPDONo].pSafety    := pMasterSafety;
        aFSoEInputPDOs[FSoEInputPDONo].pMem       := MyPara.aPara[0];
        FSoEInputPDONo += 1;
      else
        LogValue("@0490 (SafetyManager::ShareSingleConnectionInfos) Maximum limit of allowed FSoE input Frames exceeded (0x{0})", Value:=MAX_FSOE_CONNECTIONS);
      end_if;
    end_if;

    // remember that we already dealt with this connection
    pMasterConnection^.InternalConnectionState := FCS_CONNECTION;

  end_if;

END_FUNCTION

FUNCTION SafetyManager::GetObjName
	VAR_INPUT
		pThis 	: pVirtualBase;
		pTargetString 	: ^CHAR;
		TargetStringSize 	: UDINT;
	END_VAR
  VAR
  	pObjName : ^CHAR;
    ObjNameLen : UDINT;
    pEmbObjStr : ^CHAR;
    EmbObjLen : UDINT;
  END_VAR

  // check for valid this pointer
  if pThis then

    // get the name of the object
    pObjName := LSL_GetObjName(pThis);

    // check for valid name pointer
    if pObjName then
      // store the object name

      // cut the embedded object name for SCPs
      pEmbObjStr := "\SDIASSAFETYMANAGERFSOE1";
      EmbObjLen  := _strlen(src:=pEmbObjStr);
      ObjNameLen := _strlen(pObjName);
      if (ObjNameLen > EmbObjLen) & (_strcmp(str1:=pObjName + (ObjNameLen - EmbObjLen), str2:=pEmbObjStr) = 0) then
        ObjNameLen -= EmbObjLen;
      end_if;

      if ObjNameLen < TargetStringSize then
        _memcpy(pTargetString, pObjName, ObjNameLen);
        (pTargetString+ObjNameLen)^ := 0; // Insert 0 Termination
      else
        _memcpy(pTargetString, pObjName, TargetStringSize-1);
        (pTargetString + TargetStringSize-1) ^ := 0;  // Insert 0 Termination
      end_if;
    end_if;
  end_if;

END_FUNCTION

FUNCTION GLOBAL SafetyManager::SetUdpParameters
	VAR_INPUT
		pCycleTime 	: ^UDINT;
		pTimeout 	: ^UDINT;
	END_VAR

  if pCycleTime then
    sUdpVars.udOverrideCycleTime := pCycleTime^;
  end_if;

  if pTimeout then
    sUdpVars.udOverrideTimeout := pTimeout^;
  end_if;

END_FUNCTION

FUNCTION GLOBAL SafetyManager::GetUdpParameters
	VAR_INPUT
		pCycleTime 	: ^UDINT;
		pTimeout 	: ^UDINT;
	END_VAR

  if pCycleTime then
    pCycleTime^ := sUdpVars.udOverrideCycleTime;
  end_if;

  if pTimeout then
    pTimeout^ := sUdpVars.udOverrideTimeout;
  end_if;

END_FUNCTION
